// TIA Portal project "Project2" (V18)

(* hardware
DEVICE "HMI_1"  TP700 Comfort
   slot 0: "HMI_1"  TP700 Comfort  6AV2 124-0GC01-0AX0  17.0.0.0
   slot 1: "HMI_RT_1"  TP700 Comfort  6AV2 124-0GC01-0AX0  17.0.0.0
   slot 5: "HMI_1.IE_CP_1"  PROFINET Interface  17.0.0.0
      slot 1: "PROFINET Interface_1"  PROFINET Interface
         slot 1: "Port_1"  Port
         slot 2: "Port_2"  Port
   slot 7: "HMI_1.MPI/DP_CP_1"  MPI/DP Interface  17.0.0.0
DEVICE "S7-1500/ET200MP station_1"  S7-1500 station
   slot 0: "Rail_0"  Rack  6ES7 590-1***0-0AA0
   slot 1: "PLC_1"  CPU 1517-3 PN/DP  6ES7 517-3AP00-0AB0  V3.0
      slot 3: "CPU display_1"  6ES7591-1BA00-0AA0
      slot 32768: "PROFINET interface_1"  X1
         slot 32769: "Port_1"  X1 P1
         slot 32770: "Port_2"  X1 P2
      slot 33024: "PROFINET interface_2"  X2
         slot 33025: "Port_1"  X2 P1
      slot 33280: "DP interface_1"  X3
      slot 34817: "Virtual CP interface port_1"  Virtual CP interface port  Virtual CP interface port
   slot 2: "DI 16x24VDC / DQ 16x24VDC/0.5A BA_1"  DI 16x24VDC/DQ 16x24VDC/0.5A BA  6ES7 523-1BL00-0AA0  V1.1
   slot 3: "DI 16x24VDC / DQ 16x24VDC/0.5A BA_2"  DI 16x24VDC/DQ 16x24VDC/0.5A BA  6ES7 523-1BL00-0AA0  V1.1
   slot 4: "DI 16x24VDC / DQ 16x24VDC/0.5A BA_3"  DI 16x24VDC/DQ 16x24VDC/0.5A BA  6ES7 523-1BL00-0AA0  V1.1
   slot 5: "DI 16x24VDC / DQ 16x24VDC/0.5A BA_4"  DI 16x24VDC/DQ 16x24VDC/0.5A BA  6ES7 523-1BL00-0AA0  V1.1
*)

// ===== PLC "PLC_1"  CPU 1517-3 PN/DP =====

VAR_GLOBAL   // PLC tag table "Default tag table"
   "System_Byte" AT %MB1 : Byte;
   "FirstScan" AT %M1.0 : Bool;
   "DiagStatusUpdate" AT %M1.1 : Bool;
   "AlwaysTRUE" AT %M1.2 : Bool;
   "AlwaysFALSE" AT %M1.3 : Bool;
   "Clock_Byte" AT %MB0 : Byte;
   "Clock_10Hz" AT %M0.0 : Bool;
   "Clock_5Hz" AT %M0.1 : Bool;
   "Clock_2.5Hz" AT %M0.2 : Bool;
   "Clock_2Hz" AT %M0.3 : Bool;
   "Clock_1.25Hz" AT %M0.4 : Bool;
   "Clock_1Hz" AT %M0.5 : Bool;
   "Clock_0.625Hz" AT %M0.6 : Bool;
   "Clock_0.5Hz" AT %M0.7 : Bool;
END_VAR

VAR_GLOBAL   // PLC tag table "ConveyorRun_Sequence"
   "Bottle_Count" AT %MW4 : Int;
   "Start_Btn" AT %M2.0 : Bool;
   "Stop_Btn" AT %M2.1 : Bool;
   "conveyor_state" AT %M2.2 : Bool;
   "Bottle_Position" AT %MW10 : Int;
   "Clock_Edge_Mem" AT %M2.3 : Bool;
   "Crate_Count" AT %MW6 : Int;
   "Auto_State" AT %M2.4 : Bool;
   "Previous_Bottle_Count" AT %MW8 : Int;
   "Conveyor_2" AT %Q0.0 : Bool;
   "Conveyor_1" AT %Q0.1 : Bool;
END_VAR

VAR_GLOBAL   // PLC tag table "InspectionSys"
   "Fallen_Ind" AT %M8.0 : Bool;
   "EntryPE1" AT %I0.0 : Bool;
   "EntryPE2" AT %I0.1 : Bool;
   "RefreshButton" AT %M8.6 : Bool;
   "Idle_Ind" AT %M8.1 : Bool;
   "OverHeightPE_HC" AT %I0.4 : Bool;
   "TriggerPE_HC" AT %I0.2 : Bool;
   "UnderHeightPE_HC" AT %I0.3 : Bool;
   "Verifier_Okay" AT %M8.2 : Bool;
   "HCFail_Ind" AT %M8.3 : Bool;
   "HCFault_Ind" AT %M8.4 : Bool;
   "HCPass_Ind" AT %M8.5 : Bool;
   "RedLamp" AT %Q0.2 : Bool;
   "GreenLamp" AT %Q0.3 : Bool;
   "BlueLamp" AT %Q0.4 : Bool;
END_VAR

DATA_BLOCK "Inspection_Entry_DB"   // DB4
{ S7_Optimized_Access := 'TRUE' }
VERSION : 0.1
// stored: InstanceOfName Inspection_Entry
"Inspection_Entry"
BEGIN
END_DATA_BLOCK

// folder: System blocks/Program resources

DATA_BLOCK "IEC_Counter_0_DB"   // DB1
{ S7_Optimized_Access := 'TRUE' }
AUTHOR : Simatic
FAMILY : IEC
NAME : CNTR
VERSION : 1.0
// stored: InstanceOfName IEC_COUNTER
"IEC_COUNTER"
BEGIN
END_DATA_BLOCK

DATA_BLOCK "IEC_Timer_0_DB"   // DB2
{ S7_Optimized_Access := 'TRUE' }
AUTHOR : Simatic
FAMILY : IEC
NAME : IEC_TMR
VERSION : 1.0
// stored: InstanceOfName IEC_TIMER
"IEC_TIMER"
BEGIN
END_DATA_BLOCK

DATA_BLOCK "IEC_Timer_0_DB_1"   // DB3
{ S7_Optimized_Access := 'TRUE' }
AUTHOR : Simatic
FAMILY : IEC
NAME : IEC_TMR
VERSION : 1.0
// stored: InstanceOfName IEC_TIMER
"IEC_TIMER"
BEGIN
END_DATA_BLOCK

// folder: (top level)

FUNCTION_BLOCK "Inspection_Entry"   // FB1, LAD
{ S7_Optimized_Access := 'TRUE' }
VERSION : 0.1
   VAR_TEMP   // added for the SCL form of the ladder/FBD networks
      _w1 : Bool;
   END_VAR
BEGIN

REGION Network 2: Start and Stop Conveyor
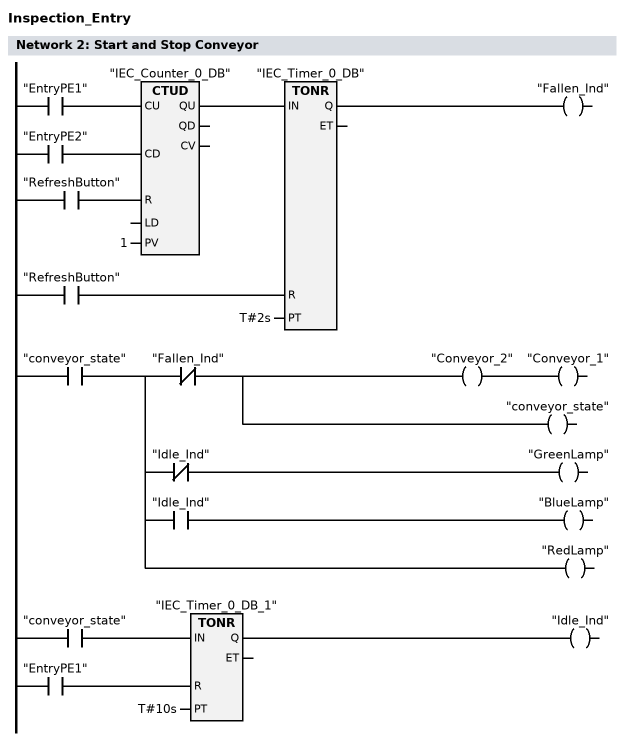
   "IEC_Counter_0_DB".CTUD(CU := "EntryPE1", CD := "EntryPE2", R := "RefreshButton", PV := 1);
   "IEC_Timer_0_DB".TONR(IN := "IEC_Counter_0_DB".QU, R := "RefreshButton", PT := T#2s);
   "Fallen_Ind" := "IEC_Timer_0_DB".Q;
   "Conveyor_2" := "conveyor_state" AND NOT "Fallen_Ind";
   "Conveyor_1" := "Conveyor_2";
   #_w1 := "conveyor_state";
   "conveyor_state" := "Conveyor_2";
   "GreenLamp" := #_w1 AND NOT "Idle_Ind";
   "BlueLamp" := #_w1 AND "Idle_Ind";
   "RedLamp" := #_w1;
   "IEC_Timer_0_DB_1".TONR(IN := "conveyor_state", R := "EntryPE1", PT := T#10s);
   "Idle_Ind" := "IEC_Timer_0_DB_1".Q;
END_REGION
END_FUNCTION_BLOCK

ORGANIZATION_BLOCK "Main"   // OB1, LAD, ProgramCycle
TITLE = "Main Program Sweep (Cycle)"
{ S7_Optimized_Access := 'TRUE' }
VERSION : 0.1
   VAR_INPUT
      Initial_Call : Bool;   // Initial call of this OB
      Remanence : Bool;   // =True, if remanent data are available
   END_VAR
   VAR_TEMP
      stop_for_man : Int;
   END_VAR
BEGIN

REGION Network 1
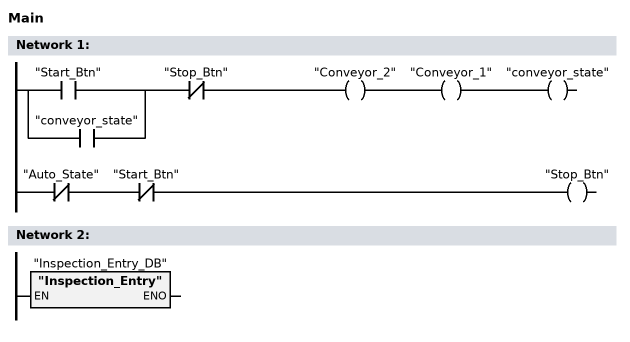
   RUNG wire#powerrail
      Contact( "Start_Btn" )
      wire#w1
      I_Contact( "Stop_Btn" )
      Coil( "Conveyor_2" )
      Coil( "Conveyor_1" )
      Coil( "conveyor_state" )
   END_RUNG
   RUNG wire#powerrail
      Contact( "conveyor_state" )
   END_RUNG wire#w1
   RUNG wire#powerrail
      I_Contact( "Auto_State" )
      I_Contact( "Start_Btn" )
      Coil( "Stop_Btn" )
   END_RUNG
   // the same network as SCL:
   "Conveyor_2" := ("Start_Btn" OR "conveyor_state") AND NOT "Stop_Btn";
   "Conveyor_1" := "Conveyor_2";
   "conveyor_state" := "Conveyor_2";
   "Stop_Btn" := NOT "Auto_State" AND NOT "Start_Btn";
END_REGION

REGION Network 2
   RUNG wire#powerrail
      "Inspection_Entry_DB"()
   END_RUNG
   // the same network as SCL:
   "Inspection_Entry_DB"();   // "Inspection_Entry"
END_REGION
END_ORGANIZATION_BLOCK

ORGANIZATION_BLOCK "Main_1"   // OB123, SCL, ProgramCycle
TITLE = "Main Program Sweep (Cycle)"
{ S7_Optimized_Access := 'TRUE' }
VERSION : 0.1
   VAR_INPUT
      Initial_Call : Bool;   // Initial call of this OB
      Remanence : Bool;   // =True, if remanent data are available
   END_VAR
BEGIN
   //TIAPortal2
   IF "conveyor_state" THEN
       // Increment position on rising edge of clock memory bit (10 Hz / 100 ms)
       IF "Clock_10Hz" AND NOT "Clock_Edge_Mem" THEN
           "Bottle_Position" := "Bottle_Position" + 10; // Step value for movement speed

           // Reset position and increment counter when bottle reaches end of belt
           IF "Bottle_Position" >= 1000 THEN
               "Bottle_Position" := 0; // Reset bottle to conveyor start
               "Previous_Bottle_Count" := "Bottle_Count";
               "Bottle_Count" := "Bottle_Count" + 1; // Increment bottle count


               IF "Bottle_Count" >= 16 THEN
                   "Bottle_Count" := 0;
                   "Crate_Count" := "Crate_Count" + 1;
               END_IF;
           END_IF;
       END_IF;
   ELSE
       "Bottle_Position" := 0; // Reset position when conveyor stops
   END_IF;

   // Update edge memory at the end of the scan (outside conveyor check)
   "Clock_Edge_Mem" := "Clock_10Hz";
END_ORGANIZATION_BLOCK

(* ===== HMI "HMI_RT_1" =====
system functions are stored by id; their names below are inferred from use
connection "HMI_Connection_1": ETHERNET, S7_1500_OMS

HMI tags "Default tag table"
   "Start_Btn" : Bool = PLC Start_Btn AT %M2.0, 1 s
   "Stop_Btn" : Bool = PLC Stop_Btn AT %M2.1, 1 s
   "conveyor_state" : Bool = PLC conveyor_state AT %M2.2, 1 s
   "Bottle_Position" : Int = PLC Bottle_Position AT %MW10, 100 ms
   "Bottle_Count" : Int = PLC Bottle_Count AT %MW4, 1 s
   "Crate_Count" : Int = PLC Crate_Count AT %MW6, 1 s
   "Auto_State" : Bool = PLC Auto_State AT %M2.4, 1 s
   "RefreshButton" : Bool = PLC RefreshButton AT %M8.6, 1 s

screen "Screen_1" 800x480
   GraphicView "Graphic view_1" at 445,151 size 354x323; Picture "Screenshot 2026-11-02 061218"
   GraphicView "Graphic view_2" at 458,410 size 65x63; Picture "Screenshot 2026-11-02 054854"
      Visibility <- "Bottle_Count"
   Button "Button_1" at 460,8 size 96x32; TextOff 'Start'
      Appearance <- "Start_Btn"
      on Press: SetBit("Start_Btn")
      on Release: ResetBit("Start_Btn")
   Button "Button_2" at 460,58 size 96x32; TextOff 'Stop'
      on Press: SetBit("Stop_Btn")
      Appearance <- "Stop_Btn"
      on Release: ResetBit("Stop_Btn")
   GraphicView "Graphic view_3" at 543,410 size 65x63; Picture "Screenshot 2026-11-02 054854"
      Visibility <- "Bottle_Count"
   GraphicView "Graphic view_4" at 632,410 size 65x63; Picture "Screenshot 2026-11-02 054854"
      Visibility <- "Bottle_Count"
   GraphicView "Graphic view_5" at 722,410 size 65x63; Picture "Screenshot 2026-11-02 054854"
      Visibility <- "Bottle_Count"
   GraphicView "Graphic view_6" at 722,330 size 65x63; Picture "Screenshot 2026-11-02 054854"
      Visibility <- "Bottle_Count"
   GraphicView "Graphic view_7" at 632,330 size 65x63; Picture "Screenshot 2026-11-02 054854"
      Visibility <- "Bottle_Count"
   GraphicView "Graphic view_8" at 542,330 size 65x63; Picture "Screenshot 2026-11-02 054854"
      Visibility <- "Bottle_Count"
   GraphicView "Graphic view_9" at 458,330 size 65x63; Picture "Screenshot 2026-11-02 054854"
      Visibility <- "Bottle_Count"
   GraphicView "Graphic view_10" at 458,250 size 65x63; Picture "Screenshot 2026-11-02 054854"
      Visibility <- "Bottle_Count"
   GraphicView "Graphic view_11" at 542,250 size 65x63; Picture "Screenshot 2026-11-02 054854"
      Visibility <- "Bottle_Count"
   GraphicView "Graphic view_12" at 635,250 size 65x63; Picture "Screenshot 2026-11-02 054854"
      Visibility <- "Bottle_Count"
   GraphicView "Graphic view_13" at 722,248 size 65x63; Picture "Screenshot 2026-11-02 054854"
      Visibility <- "Bottle_Count"
   GraphicView "Graphic view_14" at 722,171 size 65x63; Picture "Screenshot 2026-11-02 054854"
      Visibility <- "Bottle_Count"
   GraphicView "Graphic view_15" at 632,170 size 65x63; Picture "Screenshot 2026-11-02 054854"
      Visibility <- "Bottle_Count"
   GraphicView "Graphic view_16" at 542,169 size 65x63; Picture "Screenshot 2026-11-02 054854"
      Visibility <- "Bottle_Count"
   GraphicView "Graphic view_17" at 460,168 size 65x63; Picture "Screenshot 2026-11-02 054854"
      Visibility <- "Bottle_Count"
   GraphicView "Graphic view_18" at 7,280 size 45x135; Picture "Wine-bottle"
      HorizontalMovement <- "Bottle_Position"
   GraphicView "Graphic view_19" at 0,415 size 457x56; Picture "Screenshot 2026-11-02 062459"
   IOField "I/O field_1" at 604,8 size 96x32; FormatPattern s99999
      ProcessValue <- "Bottle_Count"
   Button "Button_3" at 700,8 size 96x32; TextOff 'Bottle_Cnt'
   IOField "I/O field_2" at 604,40 size 96x32; FormatPattern s99999
      ProcessValue <- "Crate_Count"
   Button "Button_4" at 697,39 size 96x32; TextOff 'Crate_Cnt'
   Switch "Switch_1" at 58,2 size 120x88; CaptionText 'Switch'; TextOff 'Man'; TextOn 'Auto'
      ProcessValue <- "Auto_State"
      on SwitchOn: SetBit("Auto_State")
      on SwitchOff: ResetBit("Auto_State")
   Button "Button_5" at 460,100 size 96x32; TextOff 'Reset'
      on Press: SetBit("RefreshButton")
      on Release: ResetBit("RefreshButton")
      Appearance <- "RefreshButton"
*)